Fanuc KAREL source: KB00029.KL

PROGRAM KB00029
%NOLOCKGROUP
%ENVIRONMENT UIF
VAR
  P1: INTEGER
  P2: STRING[80]
  P3: INTEGER
BEGIN
  P1 = 1
  P2 = 'A'
  P3 = 1
  CNC_DYN_DISI(P1, P2, P3)
END KB00029
